FUNCTION_BLOCK AUDI_FB_CTU (* Up counter (UDINT) AUDI-Adapter Version *)
  (* Standard: 61499-2; Description: Copyright (c) 2026 Meisterschulen am Ostbahnhof This program and the accompanying materials are made available under the terms of the Eclipse Public License 2.0 which is available at https://www.eclipse.org/legal/epl-2.0/ SPDX-License-Identifier: EPL-2.0 NOTE: This block fires the AX output event (Q.E1) on every update (CU, R, PV). If on-change triggering is required, use of an AX_D_FF as a filter is recommended. *)
  (* Version 1.0, 2026-04-21, Franz Höpfinger, Meisterschulen am Ostbahnhof, initial API and implementation and/or initial documentation *)
  PACKAGE adapter::iec61131::counters;
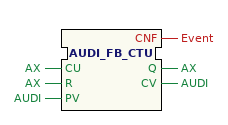
  EVENT_OUTPUT
    CNF; (* Execution Confirmation *)
  END_EVENT
  SOCKETS
    CU : adapter::types::unidirectional::AX; (* Count up *)
    R : adapter::types::unidirectional::AX; (* Reset *)
    PV : adapter::types::unidirectional::AUDI; (* Preset value *)
  END_SOCKETS
  PLUGS
    Q : adapter::types::unidirectional::AX; (* Output *)
    CV : adapter::types::unidirectional::AUDI; (* Count value *)
  END_PLUGS
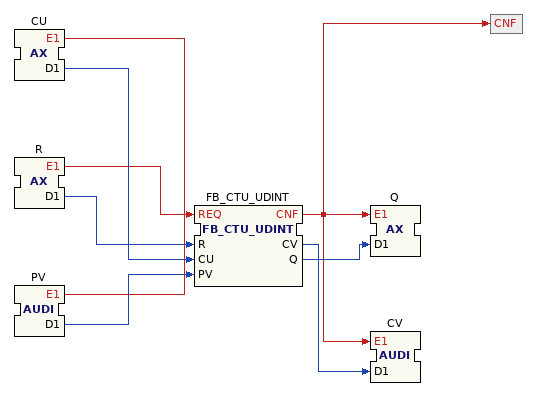
  FBS
    FB_CTU_UDINT : iec61131::counters::FB_CTU_UDINT;
  END_FBS
  EVENT_CONNECTIONS
    R.E1 TO FB_CTU_UDINT.REQ;
    CU.E1 TO FB_CTU_UDINT.REQ;
    PV.E1 TO FB_CTU_UDINT.REQ;
    FB_CTU_UDINT.CNF TO CV.E1;
    FB_CTU_UDINT.CNF TO Q.E1;
    FB_CTU_UDINT.CNF TO CNF;
  END_CONNECTIONS
  DATA_CONNECTIONS
    R.D1 TO FB_CTU_UDINT.R;
    CU.D1 TO FB_CTU_UDINT.CU;
    PV.D1 TO FB_CTU_UDINT.PV;
    FB_CTU_UDINT.CV TO CV.D1;
    FB_CTU_UDINT.Q TO Q.D1;
  END_CONNECTIONS
END_FUNCTION_BLOCK
